# EPICS substitutions: db/plsci-x86l-132.substitutions
# PLSCI records for x86l-132: FMF2, FMF3, FHF1.
# PMT numbering matches the existing all-chamber substitutions.
file "db/plsci.template"
{
    pattern { CHAMBER, PMT }
    { FMF2,1 }
    { FMF2,2 }
    { FMF2,3 }
    { FMF2,4 }
    { FMF2,5 }
    { FMF2,6 }
    { FMF2,7 }
    { FMF2,8 }
    { FMF3,1 }
    { FMF3,2 }
    { FMF3,3 }
    { FMF3,4 }
    { FMF3,5 }
    { FMF3,6 }
    { FHF1,1 }
    { FHF1,2 }
    { FHF1,3 }
    { FHF1,4 }
    { FHF1,5 }
    { FHF1,6 }
    { FHF1,7 }
    { FHF1,8 }
}
